(* IEC 61131-3 sources: plc-st-coding-agent/progress/evidence/f14_v5_public_pilot_20261112/operational_restarts/string_byte_20261112/native_probe, 2 files *)

(* ---- FB.st ---- *)
FUNCTION_BLOCK FB
VAR_OUTPUT firstByte:INT;dotByte:INT;endByte:INT;END_VAR
VAR txt:STRING(8):='1.';END_VAR
firstByte:=BYTE_TO_INT(txt[0]);dotByte:=BYTE_TO_INT(txt[1]);endByte:=BYTE_TO_INT(txt[2]);
END_FUNCTION_BLOCK

(* ---- PLC_PRG.st ---- *)
PROGRAM PLC_PRG
VAR probe:FB;step:INT;testComplete:BOOL;testPassed:BOOL:=TRUE;firstFailedStep:INT:=-1;END_VAR
IF NOT testComplete THEN
probe();
IF probe.firstByte<>49 OR probe.dotByte<>46 OR probe.endByte<>0 THEN testPassed:=FALSE;firstFailedStep:=0;END_IF;
step:=1;testComplete:=TRUE;
END_IF;
END_PROGRAM
